FUNCTION_BLOCK SimpleTest (* Simple FB with one algorithm *)
  (* Standard: 61499-1; Description: Copyright (c) 2026 Martin Erich Jobst This program and the accompanying materials are made available under the terms of the Eclipse Public License 2.0 which is available at https://www.eclipse.org/legal/epl-2.0/ SPDX-License-Identifier: EPL-2.0 *)
  (* Version 1.0, 2026-10-20, Martin Jobst *)
  {SET_ATTRIBUTE(IntegerAttribute, 6)}
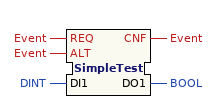
  EVENT_INPUT
    REQ; (* Normal Execution Request *)
    ALT; (* Alternate Execution Request *)
  END_EVENT
  EVENT_OUTPUT
    CNF; (* Execution Confirmation *) {SET_ATTRIBUTE(IntegerAttribute, 5)}
  END_EVENT
  VAR_INPUT
    DI1 : DINT;
  END_VAR
  VAR_OUTPUT
    DO1 : BOOL;
  END_VAR
  EC_STATES
    REQ : REQ -> CNF;
    ALT : ALT -> CNF;
  END_STATES
  ALGORITHM REQ IN ST:

  END_ALGORITHM
  ALGORITHM ALT IN ST:

  END_ALGORITHM
END_FUNCTION_BLOCK
